Fanuc KAREL source: KT00156.KL

PROGRAM KT00156
%NOLOCKGROUP
VAR
  H1: ARRAY[2] OF SHORT
  R2: REAL
  OUT: REAL
BEGIN
  H1[1] = 2
    R2 = 3.0
  OUT = H1[1] DIV R2
END KT00156
